{attribute 'qualified_only'}
VAR_GLOBAL
	
//hardware modules state linking 
//Connection-->[Message_x] Info Data
//[X] Map State
//[X] Map Diag

iModuleState1		AT %I*	:enum_FSoE_State; //104 = ok
iModuleDiag1		AT %I*	:USINT; //0 = ok
iModuleDiag1union:union_FSoE_hwDiag;


iModuleState2		AT %I*	:enum_FSoE_State;
iModuleDiag2		AT %I*	:USINT;
iModuleDiag2union:union_FSoE_hwDiag;

END_VAR

(* stored: Version 1.1.0.1, ProductVersion 3.1.4024.11
   GVL ModuleStates: Id {ab3b07d5-9ebf-0f4a-1e8d-84a72bcdb735} *)
